FUNCTION_BLOCK ToSlide (* Composite Function Block Type *)
  (* Standard: 61499-2 *)
  (* Version 0.0, 7/2/2026, template *)
  PACKAGE Main;
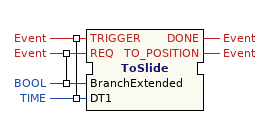
  EVENT_INPUT
    TRIGGER WITH DT1; (* Initialization Request *)
    REQ WITH BranchExtended;
  END_EVENT
  EVENT_OUTPUT
    DONE; (* Delayed Event *)
    TO_POSITION;
  END_EVENT
  VAR_INPUT
    BranchExtended : BOOL;
    DT1 : TIME; (* Delay Time *)
  END_VAR
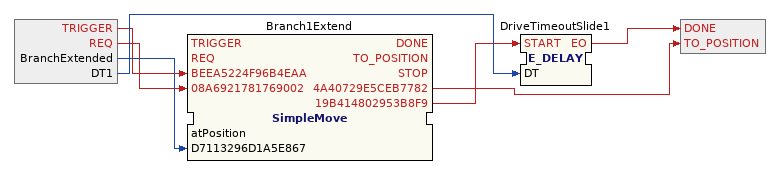
  FBS
    Branch1Extend : SimpleMove;
    DriveTimeoutSlide1 : E_DELAY;
  END_FBS
  EVENT_CONNECTIONS
    TRIGGER TO Branch1Extend.BEEA5224F96B4EAA;
    REQ TO Branch1Extend.08A6921781769002;
    Branch1Extend.4A40729E5CEB7782 TO TO_POSITION;
    DriveTimeoutSlide1.EO TO DONE;
    Branch1Extend.19B414802953B8F9 TO DriveTimeoutSlide1.START;
  END_CONNECTIONS
  DATA_CONNECTIONS
    DT1 TO DriveTimeoutSlide1.DT;
    BranchExtended TO Branch1Extend.D7113296D1A5E867;
  END_CONNECTIONS
END_FUNCTION_BLOCK
